Fanuc KAREL source: kb00154.KL

-- PROVISIONAL review KL for V770-1; original PC SHA256 a279d407ac18f4032b53814bce735154bde02d06021c74fa716f2448b2aad02e
-- Incomplete behavior may be omitted. Consult companion uncertainty JSON. Do not deploy.
PROGRAM KB00154
%NOLOCKGROUP
BEGIN
  -- UNRESOLVED_PC offsets 5-14; opcodes 3F,75
  -- UNRESOLVED_PC offsets 19-28; opcodes 3F,75
  -- UNRESOLVED_PC offsets 33-40; opcodes 9D,23
  -- UNRESOLVED_PC offsets 45-73; opcodes 27,22,2A,22,2A,22,27,9D,31
  -- UNRESOLVED_PC offsets 78-82; opcodes 7F
END KB00154
